(* IEC 61131-3 sources: Versio-VersionControlSystem/fixtures/projects/RefrigeratorControl_FBS/RefrigeratorControl.fbsproj/Device.device.xml.v3^/Plc Logic.plclogic.xml.v3^/Application.application.xml.v3^/Library/Alarm/POUs/FB_Alarm.fb.st^/Private, 6 files *)

(* ---- _M_EvaluateCommands.meth.st ---- *)
(* METADATA
{
	"v3Meta": {
		"objectGuid": "1b6999ce-aebb-4733-886d-c9adf1f6d328"
	}
}
*)
METHOD PRIVATE _M_EvaluateCommands : BOOL
// Evaluate Hmi Commands
(*IF Hmi.Cmd.Reset THEN
	// Log it
	// F_LogTrace(F_Global(Global).P_Logger, InstancePath, 'Operator Command: Reset Triggered');
	M_Reset();
END_IF*)
// Hmi.Cmd.Reset := FALSE;
END_METHOD

(* ---- _M_StateMachine.meth.st ---- *)
(* METADATA
{
	"v3Meta": {
		"objectGuid": "2939601a-39c9-43e0-ad3e-ab0b5e188b9c"
	}
}
*)
METHOD PRIVATE _M_StateMachine
// Alarm disabled
IF NOT Settings.Enable OR (NOT Condition AND State = E_AlarmState.Off) THEN
	RETURN;
END_IF

// State Machine
CASE State OF
	E_AlarmState.Off:
		IF DelayTimer.Q THEN
			NextState := E_AlarmState.Active;
		END_IF
	E_AlarmState.Active:
		IF DelayTimer.Q THEN
			NextState := E_AlarmState.Off;
		END_IF
	ELSE
		NextState := E_AlarmState.Off;
END_CASE

// Update State
_M_UpdateState();
END_METHOD

(* ---- _M_Timers.meth.st ---- *)
(* METADATA
{
	"v3Meta": {
		"objectGuid": "16b38c5d-f9c4-4a53-9840-9063bff02cb9"
	}
}
*)
METHOD PRIVATE _M_Timers : BOOL
DelayTimer.IN := SEL(State = E_AlarmState.Off, NOT (Condition OR Settings.Latch), Condition) AND Settings.Enable;
DelayTimer.PT := SEL(State = E_AlarmState.Off, Settings.OffDelayTime, Settings.OnDelayTime);
DelayTimer();
END_METHOD

(* ---- _M_UpdateState.meth.st ---- *)
(* METADATA
{
	"v3Meta": {
		"objectGuid": "97b89cef-285a-4cde-a86d-08debff8ecbf"
	}
}
*)
METHOD PRIVATE _M_UpdateState : BOOL
// Update State
IF NextState <> State THEN
	State := NextState;

	//ResetTimer
	DelayTimer(IN := FALSE);

	IF State = E_AlarmState.Off THEN
		;//Configuration.Info := '';
	END_IF
END_IF
END_METHOD

(* ---- _M_UpdateStatus.meth.st ---- *)
(* METADATA
{
	"v3Meta": {
		"objectGuid": "d2ee1933-8b70-4890-89fa-5296b2df9ef9"
	}
}
*)
METHOD PRIVATE _M_UpdateStatus : BOOL
VAR_INPUT
END_VAR

END_METHOD

(* ---- _M_EvaluateInputs.meth.st ---- *)
(* METADATA
{
	"v3Meta": {
		"objectGuid": "8322d789-b37e-4ca0-abe3-2ebac5bf988b"
	}
}
*)
METHOD PRIVATE _M_EvaluateInputs : BOOL
VAR_INST
	EnableRTrig	: R_TRIG;
	EnableFTrig	: F_TRIG;
END_VAR
// Initialized
IF Settings.ShortDesc <> '' AND NOT Configuration.Initialized THEN
	Configuration.Initialized := TRUE;
END_IF

// Enable State change
EnableRTrig(CLK := Settings.Enable);
EnableFTrig(CLK := Settings.Enable);
IF EnableRTrig.Q OR EnableFTrig.Q THEN
	NextState := E_AlarmState.Off;
	_M_UpdateState();
END_IF

// Delays
_M_Timers();
END_METHOD
